(* IEC 61131-3 sources: PortalRobot/Portal_robot/Device/application/ST/ST_AXIS_GROUP, 12 files *)

(* ---- E_AXIS_GROUP_POWER_MODE.st ---- *)
{attribute 'qualified_only'}
{attribute 'strict'}
TYPE E_AXIS_GROUP_POWER_MODE :
(
	OFF,
	OFF_REQUEST,
	ON

);
END_TYPE

(* ---- E_AXIS_GROUP_STATE.st ---- *)
{attribute 'qualified_only'}
{attribute 'strict'}
TYPE E_AXIS_GROUP_STATE :
(
	DISABLED,
	DISABLING_GROUP,
	DISABLING_POWER,
	ENABLING_POWER,
	ENABLING_GROUP,
	READY,
	MOVING_DIRECT,
	MOVING_LINEAR,
	EMG_STOP,
	HALT_STOP,
	WAIT_STOP,
	ERROR,
	RESETTING,
	RESET_VERIFY

);
END_TYPE

(* ---- E_MOTION_RESET_STATE.st ---- *)
{attribute 'qualified_only'}
{attribute 'strict'}
TYPE E_MOTION_RESET_STATE :
(
	IDLE,
	RESET_GROUP,
	WAIT_GROUP,
	RESET_AXES,
	WAIT_AXES
);
END_TYPE

(* ---- ST_AXIS_GROUP.st ---- *)
TYPE ST_AXIS_GROUP :
STRUCT
	Command     : ST_AXIS_GROUP_COMMANDS; // Команды группы осей
	Status      : ST_AXIS_GROUP_STATUS; // Рабочие статусы группы
	Diag        : ST_AXIS_GROUP_DIAGNOSTICS; // Состояние автомата и диагностика
	Error       : ST_AXIS_GROUP_ERRORS; // Активные и последние ошибки
	MotionParam : ST_AXIS_GROUP_MOTION_PARAMS; // Параметры движения
	Timeouts    : ST_AXIS_GROUP_TIMEOUTS; // Допустимое время выполнения шагов
END_STRUCT
END_TYPE

(* ---- ST_AXIS_GROUP_COMMANDS.st ---- *)
TYPE ST_AXIS_GROUP_COMMANDS :
STRUCT
	xGlobalError : BOOL; // Глобальная ошибка ячейки
	xPowerPermit : BOOL; // Разрешение включения группы при готовых физических осях
	xEnable      : BOOL; // Импульс включения группы
	xPowerEnable : BOOL; // Импульс включения группы после включения осей FB_AXIS
	xDisable     : BOOL; // Импульс отключения группы
	xReset       : BOOL; // Сброс ошибок группы
	xMoveDirect  : BOOL; // Команда прямого перемещения группы
	xMoveLinear  : BOOL; // Команда линейного перемещения группы
	xHaltCmd     : BOOL; // Команда плавной остановки
	xStopCmd     : BOOL; // Команда остановки группы
END_STRUCT
END_TYPE

(* ---- ST_AXIS_GROUP_DIAGNOSTICS.st ---- *)
TYPE ST_AXIS_GROUP_DIAGNOSTICS :
STRUCT
	iStep            : E_AXIS_GROUP_STATE; // Текущий шаг автомата группы
	iOldStep         : E_AXIS_GROUP_STATE; // Предыдущий шаг автомата
	iNewStep         : E_AXIS_GROUP_STATE; // Новый шаг после перехода
	iPowerMode       : E_AXIS_GROUP_POWER_MODE; // Текущий режим питания группы
    iLastErrorStep   : INT; // Шаг возникновения последней ошибки
    sStepName        : STRING[80]; // Текстовое имя текущего шага
    sWaitReason      : STRING[120]; // Причина ожидания на текущем шаге
    sErrorText       : STRING[120]; // Текст активной ошибки
    sWarningText     : STRING[120]; // Текст активного предупреждения
    stWarning        : ST_WARNING_EVENT; // Последнее предупреждение группы для общего журнала
    tStepPreset      : TIME; // Допустимое время текущего шага
    xStepTimeout     : BOOL; // Превышено допустимое время шага
	xStepChanged     : BOOL; // Шаг изменился в текущем цикле
    udiActualErrorID : UDINT; // Код активной ошибки
    udiLastErrorID   : UDINT; // Код последней ошибки
END_STRUCT
END_TYPE

(* ---- ST_AXIS_GROUP_ERROR.st ---- *)
TYPE ST_AXIS_GROUP_ERROR :
STRUCT
	ENABLE_ERROR          : BOOL; // Ошибка MC_GroupEnable
	POWER_ERROR           : BOOL; // Зарезервировано; питание осей контролируют FB_AXIS
	DISABLE_ERROR         : BOOL; // Ошибка MC_GroupDisable
	RESET_ERROR           : BOOL; // Ошибка MC_GroupReset
	MOVE_DIRECT_ERROR     : BOOL; // Ошибка MC_MoveDirectAbsolute
	MOVE_LINEAR_ERROR     : BOOL; // Ошибка MC_MoveLinearAbsolute
	HALT_ERROR            : BOOL; // Ошибка MC_GroupHalt
	STOP_ERROR            : BOOL; // Ошибка MC_GroupStop
	READ_POSITION_ERROR   : BOOL; // Ошибка чтения позиции группы
	READ_STATUS_ERROR     : BOOL; // Ошибка чтения статуса группы
	READ_GROUP_ERROR      : BOOL; // Ошибка чтения кода ошибки группы
	GROUP_ERROR_STOP      : BOOL; // Группа SoftMotion находится в ErrorStop
	SIMULATED_ERROR       : BOOL; // Тестовая ошибка Motion-FB, сформированная эмулятором
	OVERRIDE_ERROR        : BOOL; // Ошибка MC_GroupSetOverride
	STEP_TIMEOUT          : BOOL; // Превышено время выполнения шага
	INVALID_STATE         : BOOL; // Неизвестное состояние автомата
	POWER_PERMIT_READY    : BOOL; // Нет разрешения питания в готовности
	POWER_PERMIT_LOST     : BOOL; // Потеря разрешения питания в движении
END_STRUCT
END_TYPE

(* ---- ST_AXIS_GROUP_ERRORS.st ---- *)
TYPE ST_AXIS_GROUP_ERRORS :
STRUCT
	dwMotionErrorLatched  : DWORD; // Защёлкнутые ошибки SoftMotion
	dwLogicalErrorLatched : DWORD; // Защёлкнутые логические ошибки
	dwLogicalErrorNew     : DWORD; // Новые логические ошибки текущего цикла
	dwMotionErrorNew      : DWORD; // Новые ошибки SoftMotion текущего цикла
	dwMotionErrorActive   : DWORD; // Активные ошибки блоков SoftMotion
	dwMotionErrorPrevious : DWORD; // Ошибки SoftMotion предыдущего цикла
	dwMotionErrorLast     : DWORD; // Последняя ненулевая маска SoftMotion
	dwLogicalErrorLast    : DWORD; // Последняя ненулеевая логическая маска
	dwAlarmActive         : DWORD; // Собственные аварии группы для общего журнала
	stErrorActive         : ST_AXIS_GROUP_ERROR; // Расшифровка активных ошибок
	stErrorLast           : ST_AXIS_GROUP_ERROR; // Расшифровка последних ошибок
END_STRUCT
END_TYPE

(* ---- ST_AXIS_GROUP_FAULT_REQUEST.st ---- *)
TYPE ST_AXIS_GROUP_FAULT_REQUEST :
STRUCT
	xEnabled : BOOL; // Глобальное разрешение диагностической инъекции
	xExecute : BOOL; // Импульс формирования тестовой ошибки SM3
END_STRUCT
END_TYPE

(* ---- ST_AXIS_GROUP_MOTION_PARAMS.st ---- *)
TYPE ST_AXIS_GROUP_MOTION_PARAMS :
STRUCT
	stTargetPos      : SMC_POS_REF; // Целевая позиция в формате SoftMotion
	lrX              : LREAL := 1000; // Целевая координата X
	lrY              : LREAL := 1000; // Целевая координата Y
	lrZ              : LREAL := 1000; // Целевая координата Z
	VelFactor        : LREAL := 0.1; // Коэффициент скорости
	AccFactor        : LREAL := 0.1; // Коэффициент ускорения
	JerkFactor       : LREAL := 0.1; // Коэффициент рывка
	HaltDeceleration : LREAL := 1000; // Замедление при плавной остановке
	HaltJerk         : LREAL := 10000; // Рывок при плавной остановке
END_STRUCT
END_TYPE

(* ---- ST_AXIS_GROUP_STATUS.st ---- *)
TYPE ST_AXIS_GROUP_STATUS :
STRUCT
	xLocalError     : BOOL; // Активна любая внутренняя ошибка блока
	xLogicalError   : BOOL; // Активна логическая ошибка группы
	xGroupError     : BOOL; // Активна ошибка SoftMotion группы
	xMoveDirectDone : BOOL; // Прямое перемещение завершено
	xSimErrorAllowed: BOOL; // Разрешена безопасная тестовая инъекция ошибки SM3
	xPositionValid  : BOOL; // Координаты группы подтверждены MC_GroupReadActualPosition
	ActualX         : LREAL; // Текущая координата X
	ActualY         : LREAL; // Текущая координата Y
	ActualZ         : LREAL; // Текущая координата Z

END_STRUCT
END_TYPE

(* ---- ST_AXIS_GROUP_TIMEOUTS.st ---- *)
TYPE ST_AXIS_GROUP_TIMEOUTS :
STRUCT
    tPowerTimeout : TIME := T#5S; // Время ожидания включения или отключения питания
	tGroupTimeout : TIME := T#5S; // Время ожидания включения или отключения группы
    tStopTimeout  : TIME := T#5S; // Время ожидания остановки
	tHaltTimeout  : TIME := T#5S; // Время ожидания плавной остановки
    tHomeTimeout  : TIME := T#30S; // Время ожидания поиска домашней позиции
    tMoveTimeout  : TIME := T#30S; // Время ожидания завершения перемещения
END_STRUCT
END_TYPE
